SUBAPPLICATION ALI_GT_0 (* Prüft ob LINT-Adapter Wert > 0 ist (AX-Adapter Ausgang) *)
  (* Standard: 61499-2 *)
  (* Version 1.0, 2026-10-15, franz, Meisterschulen am Ostbahnhof *)
  PACKAGE MyLib::sys;
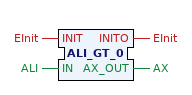
  EVENT_INPUT
    INIT : EInit; (* Initialization Request *)
  END_EVENT
  EVENT_OUTPUT
    INITO : EInit; (* Initialization Confirm *)
  END_EVENT
  SOCKETS
    IN : adapter::types::unidirectional::ALI;
  END_SOCKETS
  PLUGS
    AX_OUT : adapter::types::unidirectional::AX;
  END_PLUGS
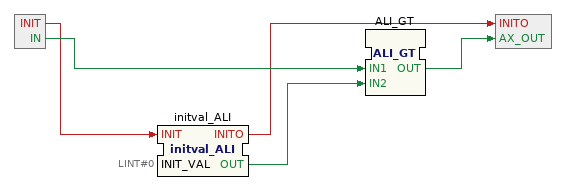
  FBS
    ALI_GT : adapter::iec61131::comparison::ALI_GT;
    initval_ALI : adapter::types::unidirectional::ALI::initval::initval_ALI(INIT_VAL := LINT#0);
  END_FBS
  EVENT_CONNECTIONS
    INIT TO initval_ALI.INIT;
    initval_ALI.INITO TO INITO;
  END_CONNECTIONS
  ADAPTER_CONNECTIONS
    IN TO ALI_GT.IN1;
    ALI_GT.OUT TO AX_OUT;
    initval_ALI.OUT TO ALI_GT.IN2;
  END_CONNECTIONS
END_SUBAPPLICATION
